Fanuc KAREL source: kf00045.KL

-- PROVISIONAL review KL for V1013-1; original PC SHA256 a82d14f3ccf68cbebacd881832450efd4e4816f861ff26c19c1a8e190ca08fb8
-- Incomplete behavior may be omitted. Consult companion uncertainty JSON. Do not deploy.
PROGRAM KF00045
%NOLOCKGROUP
VAR
  I : INTEGER
  J : INTEGER
  X : REAL
  Y : REAL
  B : BOOLEAN
  C : BOOLEAN
  TXT : STRING[80]
  TXT2 : STRING[80]
  STATUS : INTEGER
-- UNRESOLVED_DECL AI type=002010
-- UNRESOLVED_DECL BI type=002010
-- UNRESOLVED_DECL P type=000102
-- UNRESOLVED_DECL JP type=000199
-- UNRESOLVED_DECL PF type=000101
-- UNRESOLVED_DECL V1 type=000013
-- UNRESOLVED_DECL V2 type=000013
BEGIN
  -- UNRESOLVED_PC offsets 5-12; opcodes 9D,23
  -- UNRESOLVED_PC offsets 17-30; opcodes 21,9D,57,79
  -- UNRESOLVED_PC offsets 35-49; opcodes 21,9D,52,23
  -- UNRESOLVED_PC offsets 59-63; opcodes 7F
END KF00045
